(* Logix 5000 project; controller R400_500_XLS vendor 1 type 14 code 216 rev 31.11; software revision 31.01; part 21 of 32 *)
(* tags used below, declared in another part *)
   Abort1 : DINT;   // Not Used
   Alarm : SINT;   // Wait 3 seconds
   AlarmAcked : BOOL;   // Alarm has been acked
   bAlrm : BOOL[64];
   CycExcBuffer : UDT_CYCLE;
   F1rinse : DINT;   // Not Used
   F3rinse : DINT;   // Not Used
   H0_Temp : REAL;
   H1_Temp : REAL;
   HDelta_T : REAL;
   HeatSmp : DINT;
   iBuffer : DINT[5];
   Inj_Cond : SINT;   // Conductivity injection based steps
   Last_Hdelta_T : REAL;
   M : DINT[5];   // Memory Bits
   ONS_FC01 : DINT;
   ONS_FC12 : DINT;
   PresetMin : SINT;
   PresetSec : SINT;
   PreWtrDrnTme : DINT;
   PwExcBuffer : UDT_PW;
   PWR_UP : DINT;
   rBuffer : REAL[4];
   RecircLowHysteresis : REAL;
   RinseExcBuffer : UDT_RINSE;
   Run : DINT;
   SmpDrnTme : DINT;
   SmpHeatingSp : REAL;
   SmpLowHysteresis : REAL;
   StartPump3 : BOOL;   // Main Pump running
   Tmr : TIMER[107];
   TrecircSec : DINT;
   Trt_PrWsh : DINT;
   Trt_Rinse : DINT;   // Rinse steps
   washerMode : SINT;   // Washer Mode Flag 0 -> Ready; 1 -> Supervisor; 2 -> Service; 3 -> Run.
   WSH56_StartHeating : BOOL;   // Start heating
   WSH56_StartRecirculation : BOOL;   // Start the recirculation
   WshExcBuffer : UDT_WASH;
   Cfg_10_Modules : BOOL;   // Chassis is configured 10 slots
   Cfg_11_Modules : BOOL;
   Ctrlr_Status : DINT;
   Current_Screen : DINT;
   I_Ld_Dr_Cls_Sw : BOOL;   // Load door close
   I_MCR : BOOL;   // MCR input
   I_Pw_Tnk_Lvl_Sw : BOOL;   // Pure water tank level switch
   I_Smp_Lvl_Hgh : BOOL;   // Sump high level switch
   I_Smp_Lvl_Lw : BOOL;   // Sump low level switch
   I_Unld_Dr_Cls_Sw : BOOL;   // Unload door close
   MaintainCloseLd : BOOL;
   MaintainCloseUnld : BOOL;
   msg : BOOL[512];
   Msg_PwrUp : DINT;
   s007 : DINT;
   Screen_Ctrl : DINT;   // PLC Screen Request
   SumpHeatAlmRate : REAL;
   SumpTemp : REAL;   // Sump temperature in °C
   Unit : Hrdwre;   // Unit Configuration
(* MainProgram, continued *)

ROUTINE WSH_12_PWR_UP   (* ladder *)
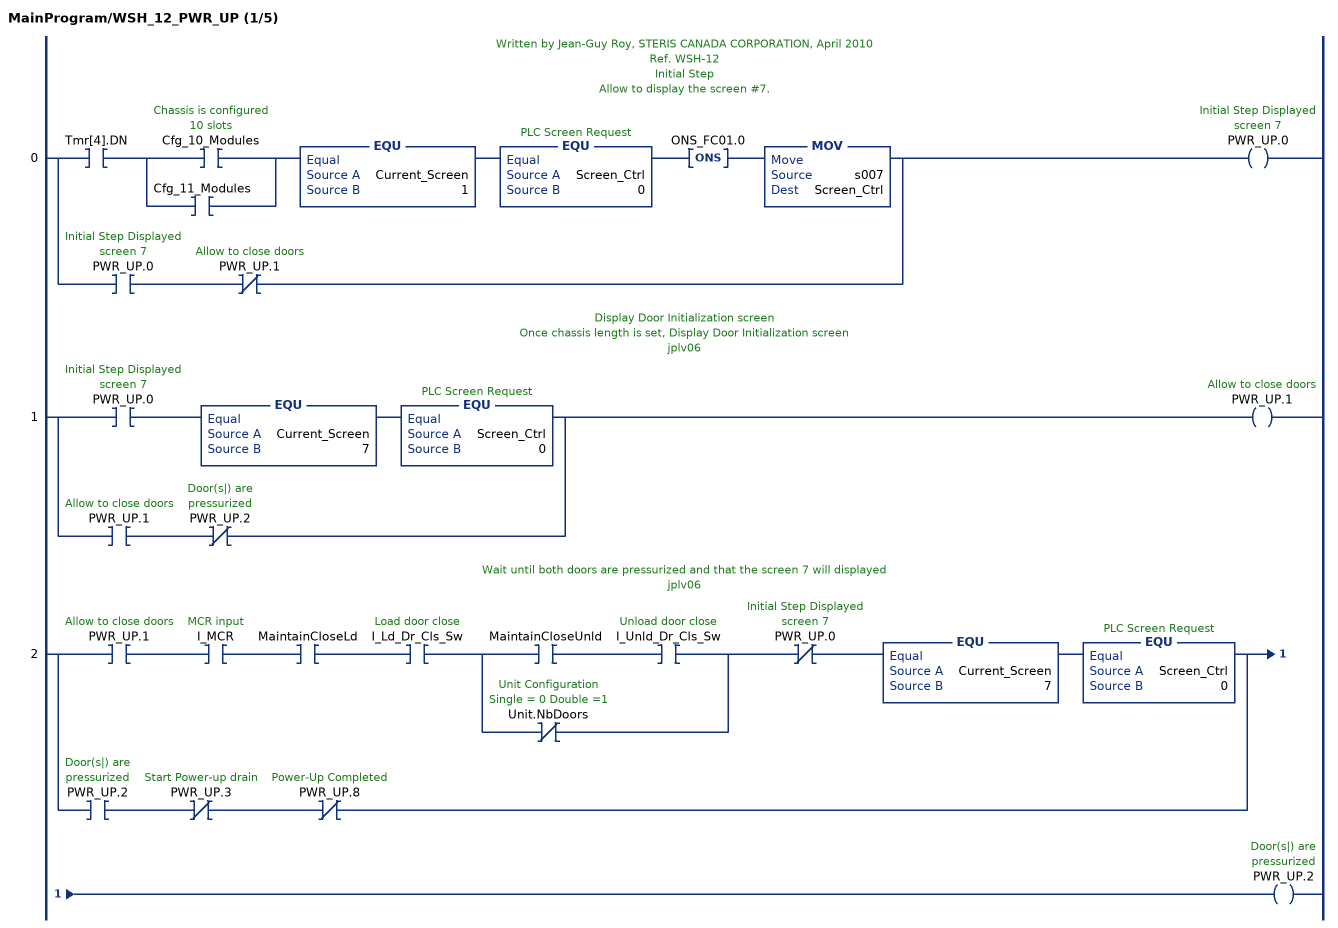
   // Written by Jean-Guy Roy, STERIS CANADA CORPORATION, April 2010
   // Ref. WSH-12
   // Initial Step
   // Allow to display the screen #7.
   0: [XIC(Tmr[4].DN) [XIC(Cfg_10_Modules) ,XIC(Cfg_11_Modules) ] EQU(Current_Screen,1) EQU(Screen_Ctrl,0) ONS(ONS_FC01.0) MOV(s007,Screen_Ctrl) ,XIC(PWR_UP.0) XIO(PWR_UP.1) ]OTE(PWR_UP.0);
   // Display Door Initialization screen
   // Once chassis length is set, Display Door Initialization screen
   // jplv06
   1: [XIC(PWR_UP.0) EQU(Current_Screen,7) EQU(Screen_Ctrl,0) ,XIC(PWR_UP.1) XIO(PWR_UP.2) ]OTE(PWR_UP.1);
   // Wait until both doors are pressurized and that the screen 7 will displayed
   // jplv06
   2: [XIC(PWR_UP.1) XIC(I_MCR) XIC(MaintainCloseLd) XIC(I_Ld_Dr_Cls_Sw) [XIC(MaintainCloseUnld) XIC(I_Unld_Dr_Cls_Sw) ,XIO(Unit.NbDoors) ] XIO(PWR_UP.0) EQU(Current_Screen,7) EQU(Screen_Ctrl,0) ,XIC(PWR_UP.2) XIO(PWR_UP.3) XIO(PWR_UP.8) ]OTE(PWR_UP.2);
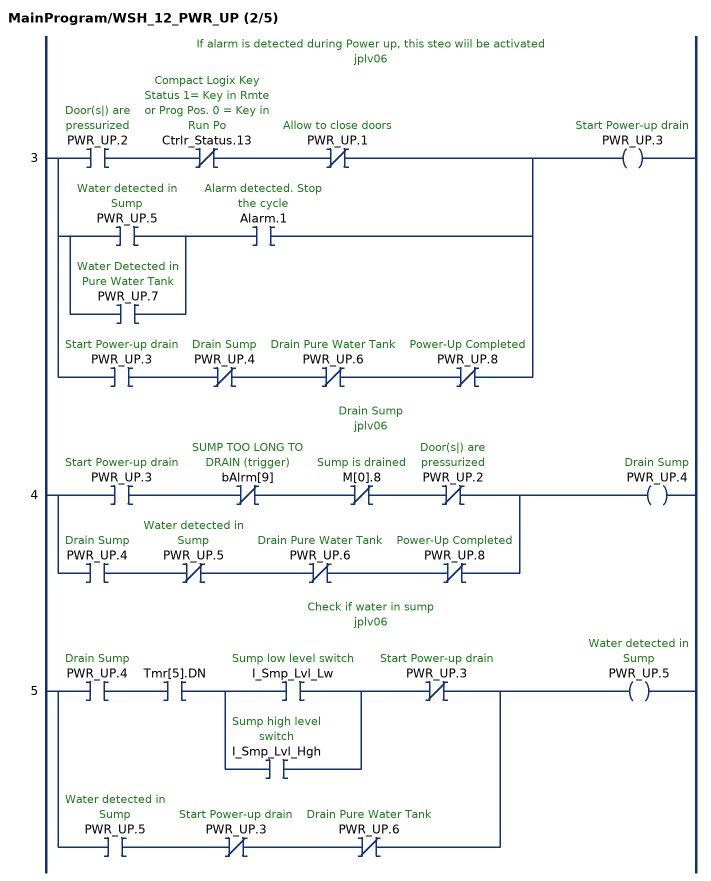
   // If alarm is detected during Power up, this steo wiil be activated
   // jplv06
   3: [XIC(PWR_UP.2) XIO(Ctrlr_Status.13) XIO(PWR_UP.1) ,[XIC(PWR_UP.5) ,XIC(PWR_UP.7) ] XIC(Alarm.1) ,XIC(PWR_UP.3) XIO(PWR_UP.4) XIO(PWR_UP.6) XIO(PWR_UP.8) ]OTE(PWR_UP.3);
   // Drain Sump
   // jplv06
   4: [XIC(PWR_UP.3) XIO(bAlrm[9]) XIO(M[0].8) XIO(PWR_UP.2) ,XIC(PWR_UP.4) XIO(PWR_UP.5) XIO(PWR_UP.6) XIO(PWR_UP.8) ]OTE(PWR_UP.4);
   // Check if water in sump
   // jplv06
   5: [XIC(PWR_UP.4) XIC(Tmr[5].DN) [XIC(I_Smp_Lvl_Lw) ,XIC(I_Smp_Lvl_Hgh) ] XIO(PWR_UP.3) ,XIC(PWR_UP.5) XIO(PWR_UP.3) XIO(PWR_UP.6) ]OTE(PWR_UP.5);
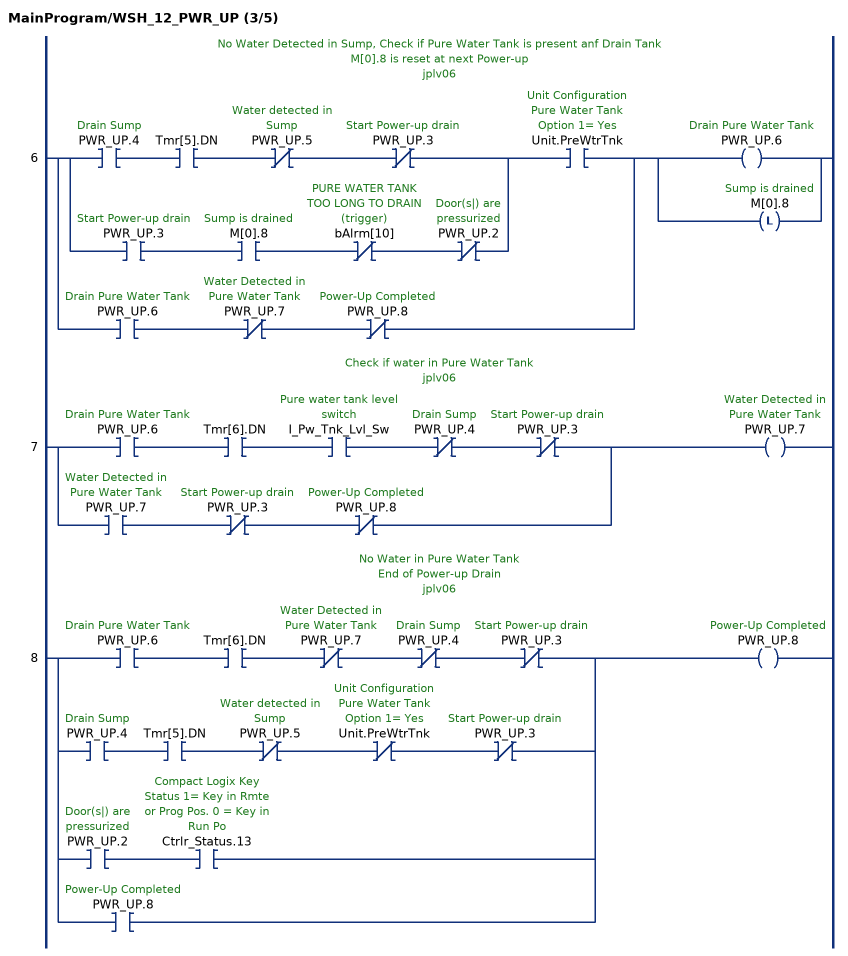
   // No Water Detected in Sump, Check if Pure Water Tank is present anf Drain Tank
   // M[0].8 is reset at next Power-up
   // jplv06
   6: [[XIC(PWR_UP.4) XIC(Tmr[5].DN) XIO(PWR_UP.5) XIO(PWR_UP.3) ,XIC(PWR_UP.3) XIC(M[0].8) XIO(bAlrm[10]) XIO(PWR_UP.2) ] XIC(Unit.PreWtrTnk) ,XIC(PWR_UP.6) XIO(PWR_UP.7) XIO(PWR_UP.8) ][OTE(PWR_UP.6) ,OTL(M[0].8) ];
   // Check if water in Pure Water Tank
   // jplv06
   7: [XIC(PWR_UP.6) XIC(Tmr[6].DN) XIC(I_Pw_Tnk_Lvl_Sw) XIO(PWR_UP.4) XIO(PWR_UP.3) ,XIC(PWR_UP.7) XIO(PWR_UP.3) XIO(PWR_UP.8) ]OTE(PWR_UP.7);
   // No Water in Pure Water Tank
   // End of Power-up Drain
   // jplv06
   8: [[XIC(PWR_UP.6) XIC(Tmr[6].DN) XIO(PWR_UP.7) XIO(PWR_UP.4) XIO(PWR_UP.3) ,XIC(PWR_UP.4) XIC(Tmr[5].DN) XIO(PWR_UP.5) XIO(Unit.PreWtrTnk) XIO(PWR_UP.3) ,XIC(PWR_UP.2) XIC(Ctrlr_Status.13) ] ,XIC(PWR_UP.8) ]OTE(PWR_UP.8);
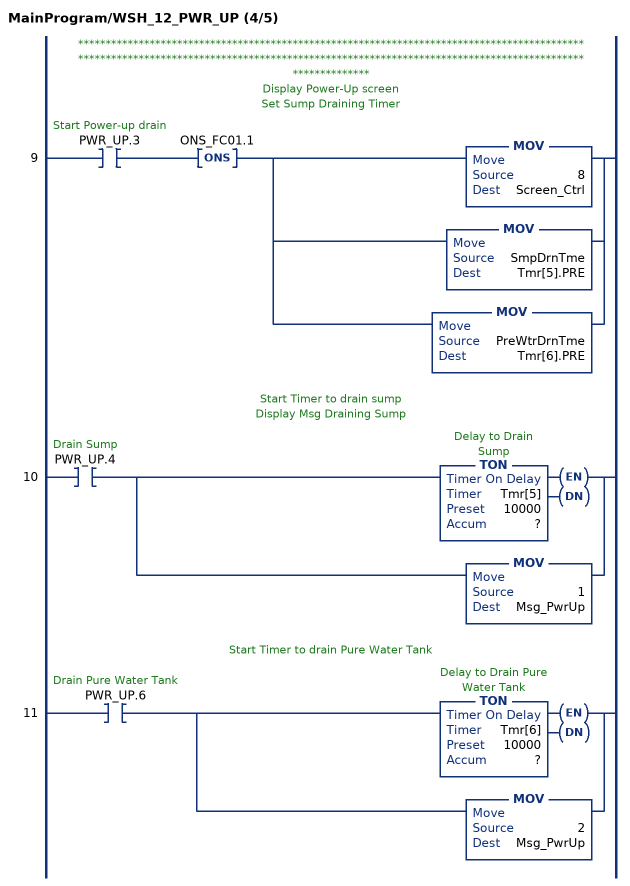
   // ******************************************************************************************************************************************************************************************************
   // Display Power-Up screen
   // Set Sump Draining Timer
   9: XIC(PWR_UP.3)ONS(ONS_FC01.1)[MOV(8,Screen_Ctrl) ,MOV(SmpDrnTme,Tmr[5].PRE) ,MOV(PreWtrDrnTme,Tmr[6].PRE) ];
   // Start Timer to drain sump
   // Display Msg Draining Sump
   10: XIC(PWR_UP.4)[TON(Tmr[5],?,?) ,MOV(1,Msg_PwrUp) ];
   // Start Timer to drain Pure Water Tank
   11: XIC(PWR_UP.6)[TON(Tmr[6],?,?) ,MOV(2,Msg_PwrUp) ];
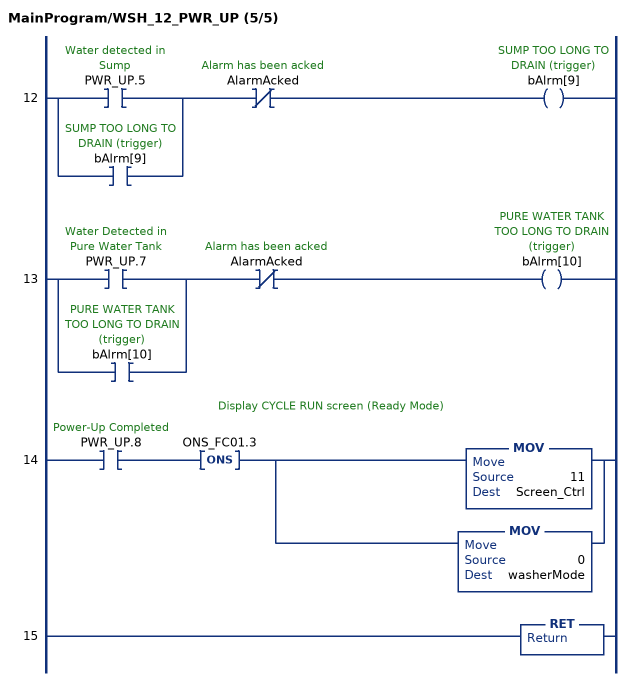
   12: [XIC(PWR_UP.5) ,XIC(bAlrm[9]) ]XIO(AlarmAcked)OTE(bAlrm[9]);
   13: [XIC(PWR_UP.7) ,XIC(bAlrm[10]) ]XIO(AlarmAcked)OTE(bAlrm[10]);
   // Display CYCLE RUN screen (Ready Mode)
   14: XIC(PWR_UP.8)ONS(ONS_FC01.3)[MOV(11,Screen_Ctrl) ,MOV(0,washerMode) ];
   15: RET();
END_ROUTINE

ROUTINE WSH_15_WSH_31_RECIRC_HEAT_SUMP   (* ladder *)
// This module is to heat the sump and the control of the recirculation timer
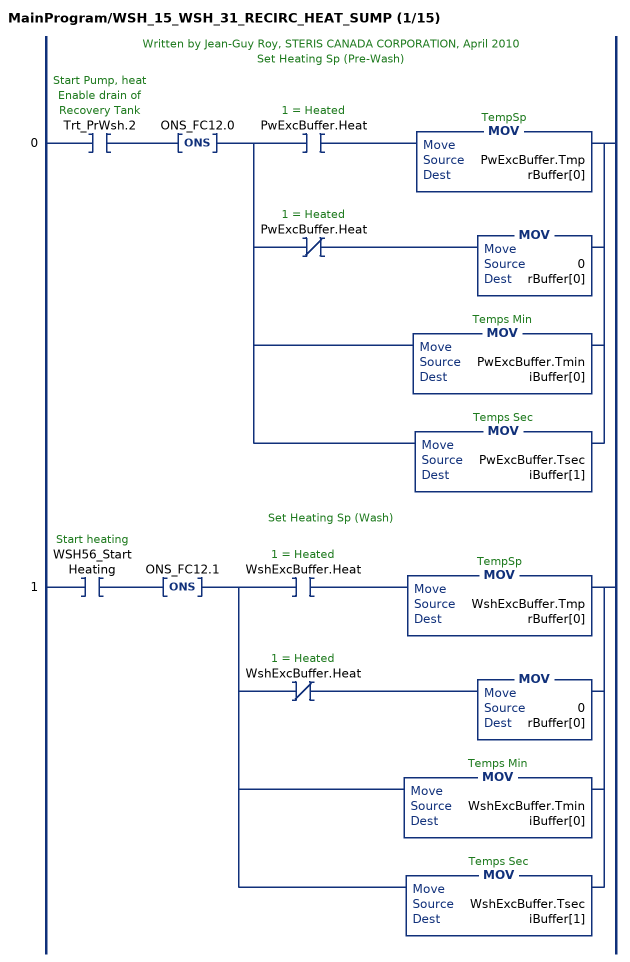
   // Written by Jean-Guy Roy, STERIS CANADA CORPORATION, April 2010
   // Set Heating Sp (Pre-Wash)
   0: XIC(Trt_PrWsh.2)ONS(ONS_FC12.0)[XIC(PwExcBuffer.Heat) MOV(PwExcBuffer.Tmp,rBuffer[0]) ,XIO(PwExcBuffer.Heat) MOV(0,rBuffer[0]) ,MOV(PwExcBuffer.Tmin,iBuffer[0]) ,MOV(PwExcBuffer.Tsec,iBuffer[1]) ];
   // Set Heating Sp (Wash)
   1: XIC(WSH56_StartHeating)ONS(ONS_FC12.1)[XIC(WshExcBuffer.Heat) MOV(WshExcBuffer.Tmp,rBuffer[0]) ,XIO(WshExcBuffer.Heat) MOV(0,rBuffer[0]) ,MOV(WshExcBuffer.Tmin,iBuffer[0]) ,MOV(WshExcBuffer.Tsec,iBuffer[1]) ];
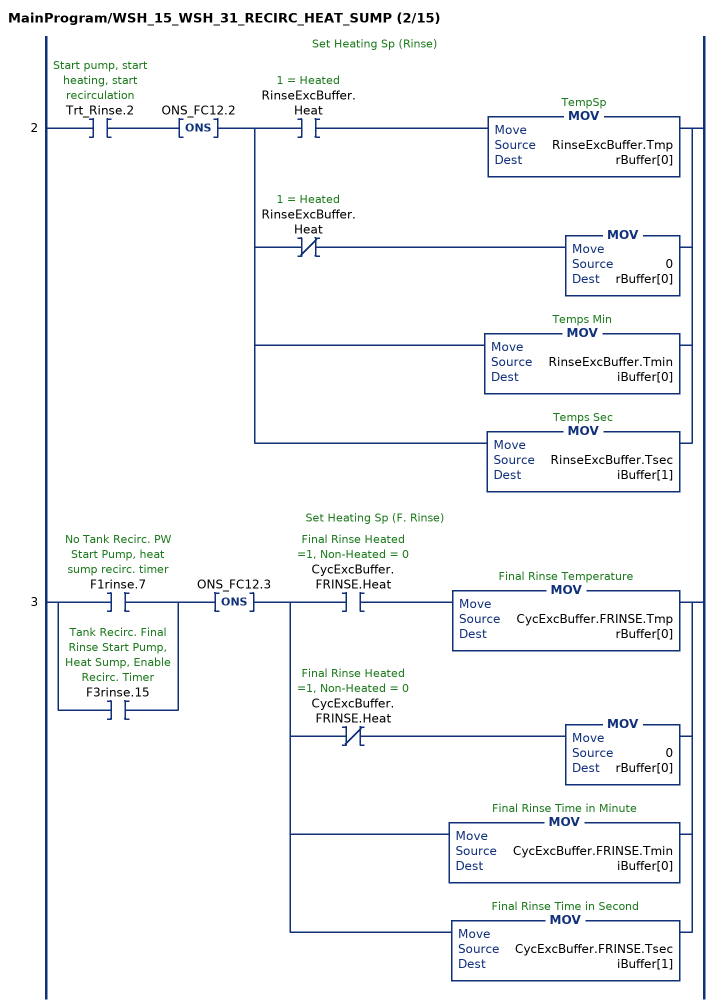
   // Set Heating Sp (Rinse)
   2: XIC(Trt_Rinse.2)ONS(ONS_FC12.2)[XIC(RinseExcBuffer.Heat) MOV(RinseExcBuffer.Tmp,rBuffer[0]) ,XIO(RinseExcBuffer.Heat) MOV(0,rBuffer[0]) ,MOV(RinseExcBuffer.Tmin,iBuffer[0]) ,MOV(RinseExcBuffer.Tsec,iBuffer[1]) ];
   // Set Heating Sp (F. Rinse)
   3: [XIC(F1rinse.7) ,XIC(F3rinse.15) ]ONS(ONS_FC12.3)[XIC(CycExcBuffer.FRINSE.Heat) MOV(CycExcBuffer.FRINSE.Tmp,rBuffer[0]) ,XIO(CycExcBuffer.FRINSE.Heat) MOV(0,rBuffer[0]) ,MOV(CycExcBuffer.FRINSE.Tmin,iBuffer[0]) ,MOV(CycExcBuffer.FRINSE.Tsec,iBuffer[1]) ];
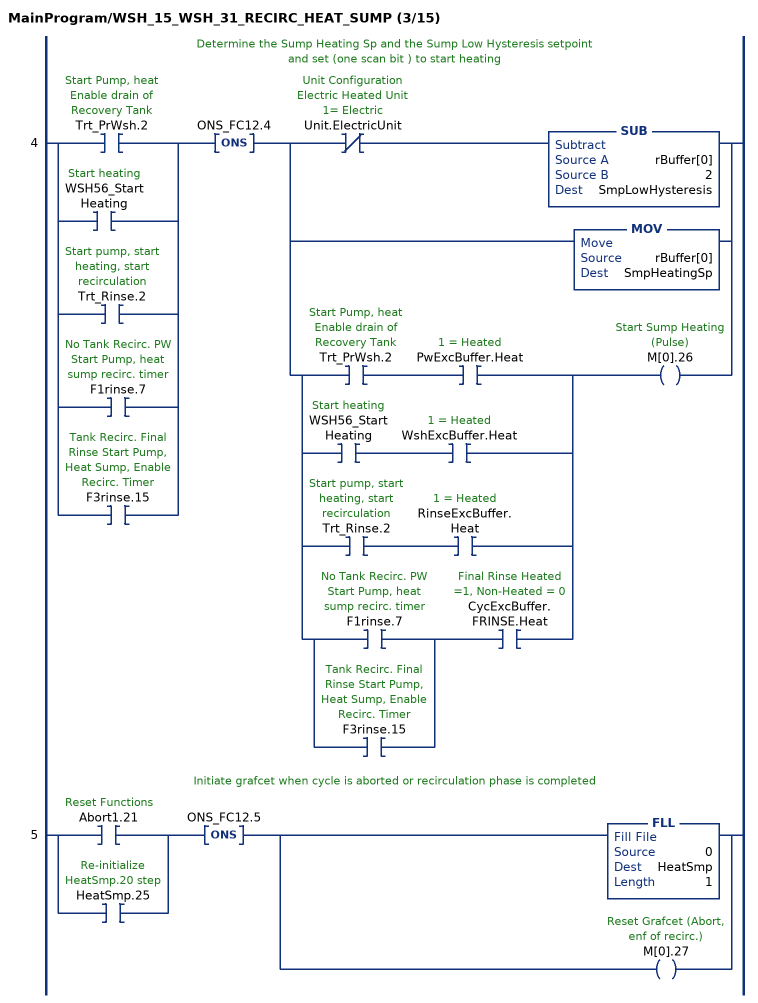
   // Determine the Sump Heating Sp and the Sump Low Hysteresis setpoint
   // and set (one scan bit ) to start heating
   4: [XIC(Trt_PrWsh.2) ,XIC(WSH56_StartHeating) ,XIC(Trt_Rinse.2) ,XIC(F1rinse.7) ,XIC(F3rinse.15) ]ONS(ONS_FC12.4)[XIO(Unit.ElectricUnit) SUB(rBuffer[0],2,SmpLowHysteresis) ,MOV(rBuffer[0],SmpHeatingSp) ,[XIC(Trt_PrWsh.2) XIC(PwExcBuffer.Heat) ,XIC(WSH56_StartHeating) XIC(WshExcBuffer.Heat) ,XIC(Trt_Rinse.2) XIC(RinseExcBuffer.Heat) ,[XIC(F1rinse.7) ,XIC(F3rinse.15) ] XIC(CycExcBuffer.FRINSE.Heat) ] OTE(M[0].26) ];
   // Initiate grafcet when cycle is aborted or recirculation phase is completed
   5: [XIC(Abort1.21) ,XIC(HeatSmp.25) ]ONS(ONS_FC12.5)[FLL(0,HeatSmp,1) ,OTE(M[0].27) ];
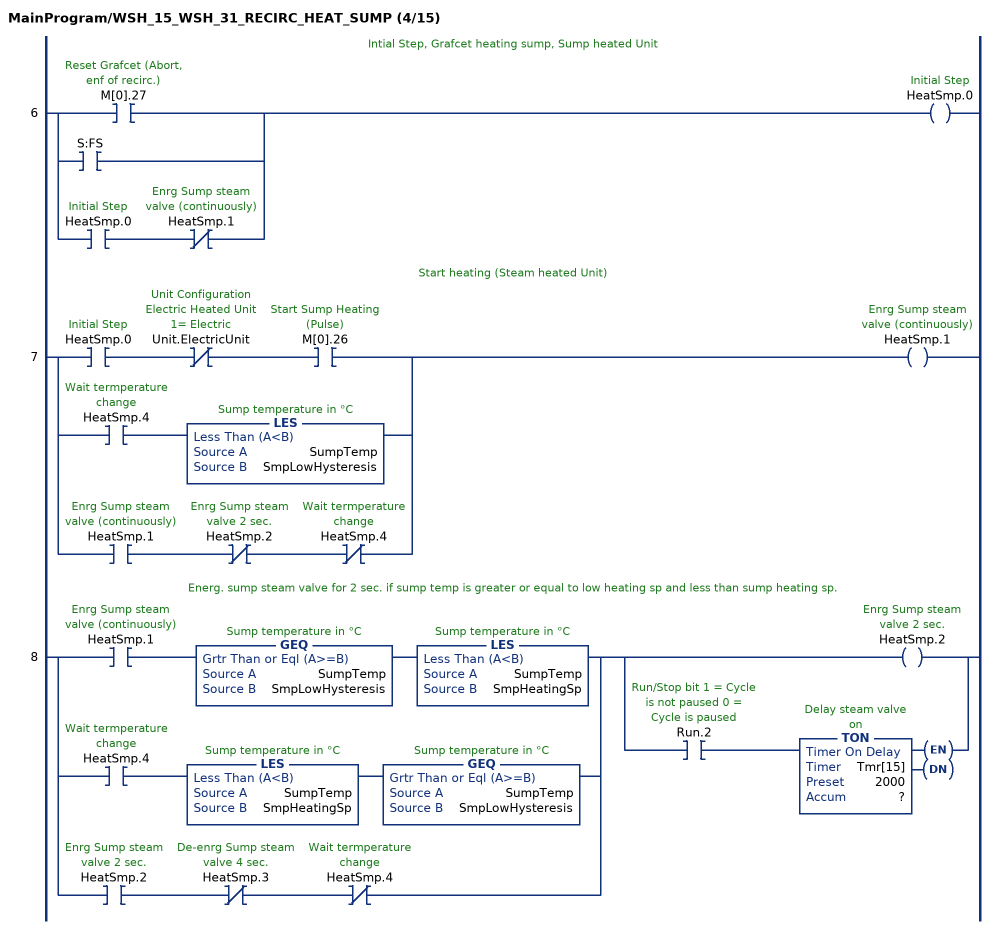
   // Intial Step, Grafcet heating sump, Sump heated Unit
   6: [XIC(M[0].27) ,XIC(S:FS) ,XIC(HeatSmp.0) XIO(HeatSmp.1) ]OTE(HeatSmp.0);
   // Start heating (Steam heated Unit)
   7: [XIC(HeatSmp.0) XIO(Unit.ElectricUnit) XIC(M[0].26) ,XIC(HeatSmp.4) LES(SumpTemp,SmpLowHysteresis) ,XIC(HeatSmp.1) XIO(HeatSmp.2) XIO(HeatSmp.4) ]OTE(HeatSmp.1);
   // Energ. sump steam valve for 2 sec. if sump temp is greater or equal to low heating sp and less than sump heating sp.
   8: [XIC(HeatSmp.1) GEQ(SumpTemp,SmpLowHysteresis) LES(SumpTemp,SmpHeatingSp) ,XIC(HeatSmp.4) LES(SumpTemp,SmpHeatingSp) GEQ(SumpTemp,SmpLowHysteresis) ,XIC(HeatSmp.2) XIO(HeatSmp.3) XIO(HeatSmp.4) ][OTE(HeatSmp.2) ,XIC(Run.2) TON(Tmr[15],?,?) ];
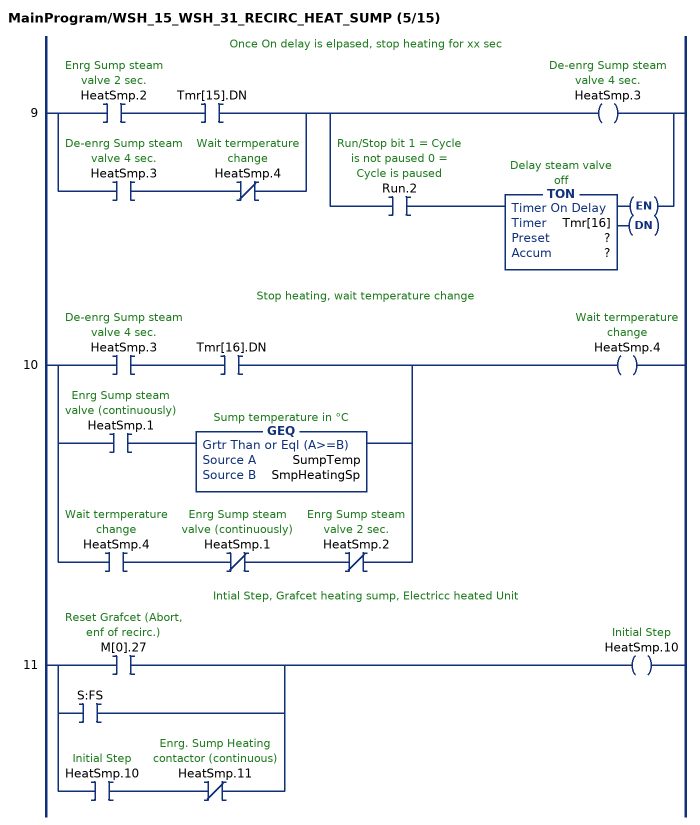
   // Once On delay is elpased, stop heating for xx sec
   9: [XIC(HeatSmp.2) XIC(Tmr[15].DN) ,XIC(HeatSmp.3) XIO(HeatSmp.4) ][OTE(HeatSmp.3) ,XIC(Run.2) TON(Tmr[16],?,?) ];
   // Stop heating, wait temperature change
   10: [XIC(HeatSmp.3) XIC(Tmr[16].DN) ,XIC(HeatSmp.1) GEQ(SumpTemp,SmpHeatingSp) ,XIC(HeatSmp.4) XIO(HeatSmp.1) XIO(HeatSmp.2) ]OTE(HeatSmp.4);
   // Intial Step, Grafcet heating sump, Electricc heated Unit
   11: [XIC(M[0].27) ,XIC(S:FS) ,XIC(HeatSmp.10) XIO(HeatSmp.11) ]OTE(HeatSmp.10);
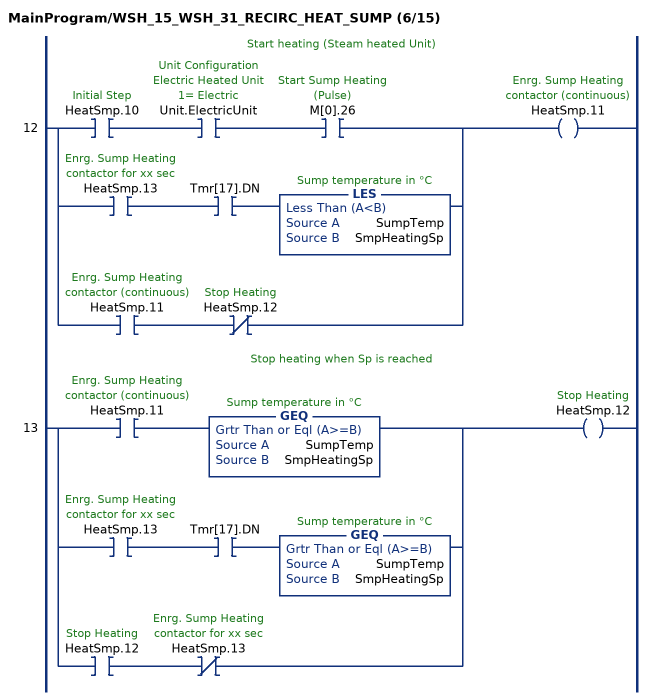
   // Start heating (Steam heated Unit)
   12: [XIC(HeatSmp.10) XIC(Unit.ElectricUnit) XIC(M[0].26) ,XIC(HeatSmp.13) XIC(Tmr[17].DN) LES(SumpTemp,SmpHeatingSp) ,XIC(HeatSmp.11) XIO(HeatSmp.12) ]OTE(HeatSmp.11);
   // Stop heating when Sp is reached
   13: [XIC(HeatSmp.11) GEQ(SumpTemp,SmpHeatingSp) ,XIC(HeatSmp.13) XIC(Tmr[17].DN) GEQ(SumpTemp,SmpHeatingSp) ,XIC(HeatSmp.12) XIO(HeatSmp.13) ]OTE(HeatSmp.12);
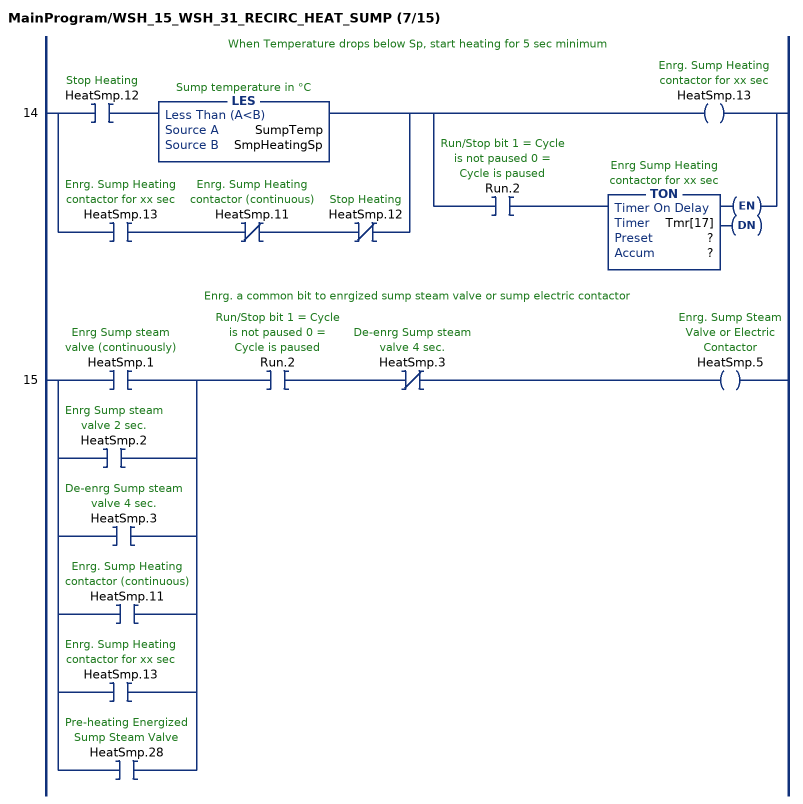
   // When Temperature drops below Sp, start heating for 5 sec minimum
   14: [XIC(HeatSmp.12) LES(SumpTemp,SmpHeatingSp) ,XIC(HeatSmp.13) XIO(HeatSmp.11) XIO(HeatSmp.12) ][OTE(HeatSmp.13) ,XIC(Run.2) TON(Tmr[17],?,?) ];
   // Enrg. a common bit to enrgized sump steam valve or sump electric contactor
   15: [XIC(HeatSmp.1) ,XIC(HeatSmp.2) ,XIC(HeatSmp.3) ,XIC(HeatSmp.11) ,XIC(HeatSmp.13) ,XIC(HeatSmp.28) ]XIC(Run.2)XIO(HeatSmp.3)OTE(HeatSmp.5);
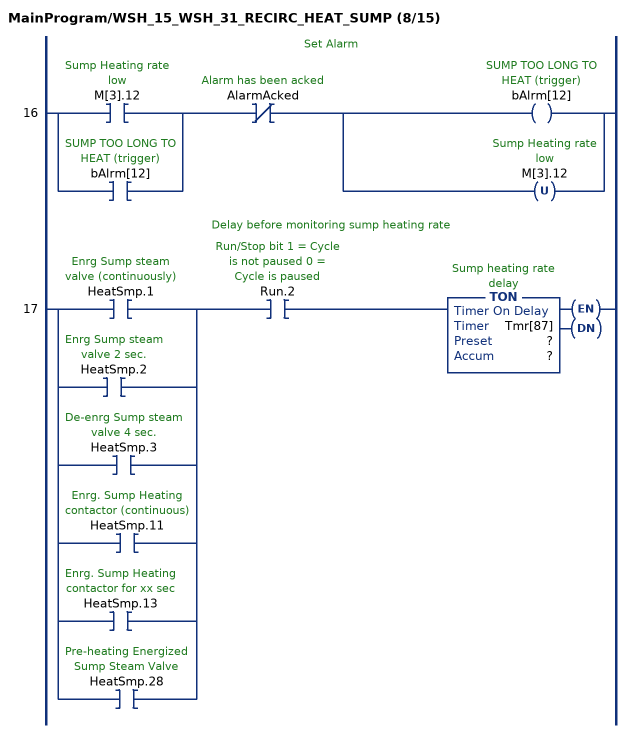
   // Set Alarm
   16: [XIC(M[3].12) ,XIC(bAlrm[12]) ]XIO(AlarmAcked)[OTE(bAlrm[12]) ,OTU(M[3].12) ];
   // Delay before monitoring sump heating rate
   17: [XIC(HeatSmp.1) ,XIC(HeatSmp.2) ,XIC(HeatSmp.3) ,XIC(HeatSmp.11) ,XIC(HeatSmp.13) ,XIC(HeatSmp.28) ]XIC(Run.2)TON(Tmr[87],?,?);
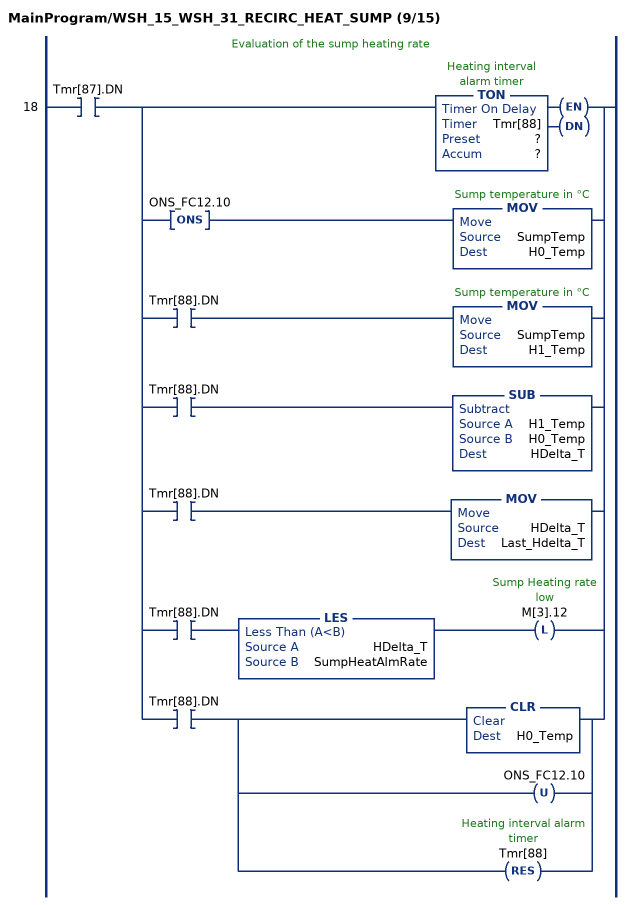
   // Evaluation of the sump heating rate
   18: XIC(Tmr[87].DN)[TON(Tmr[88],?,?) ,ONS(ONS_FC12.10) MOV(SumpTemp,H0_Temp) ,XIC(Tmr[88].DN) MOV(SumpTemp,H1_Temp) ,XIC(Tmr[88].DN) SUB(H1_Temp,H0_Temp,HDelta_T) ,XIC(Tmr[88].DN) MOV(HDelta_T,Last_Hdelta_T) ,XIC(Tmr[88].DN) LES(HDelta_T,SumpHeatAlmRate) OTL(M[3].12) ,XIC(Tmr[88].DN) [CLR(H0_Temp) ,OTU(ONS_FC12.10) ,RES(Tmr[88]) ] ];
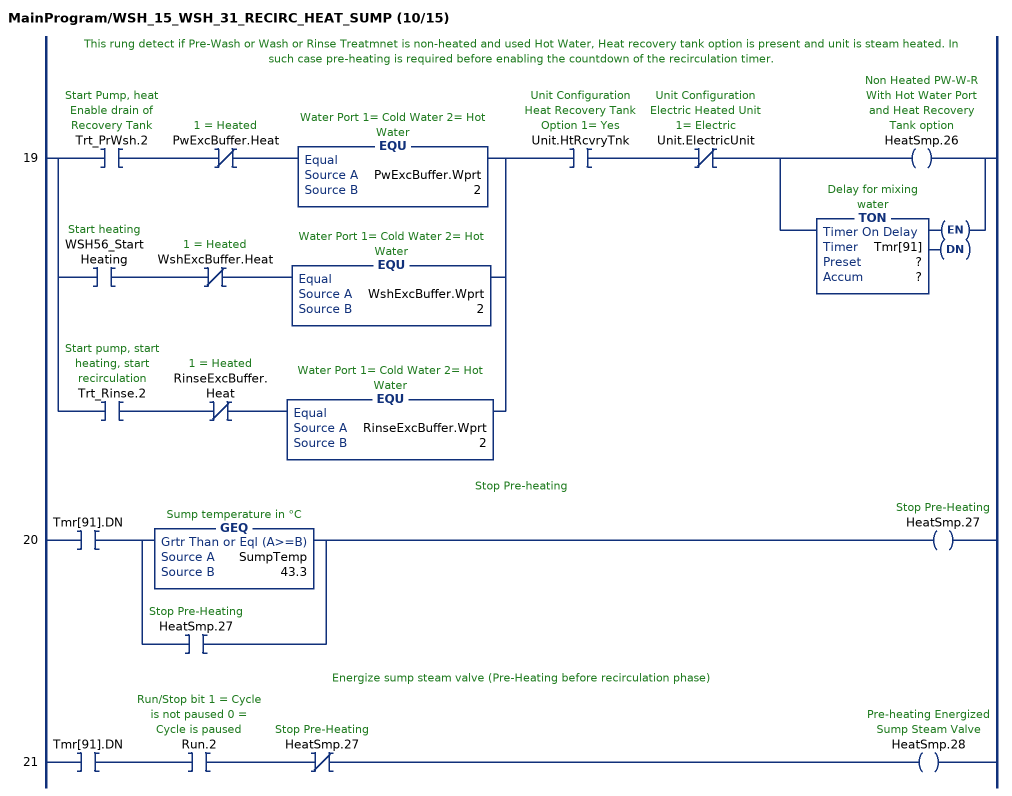
   // This rung detect if Pre-Wash or Wash or Rinse Treatmnet is non-heated and used Hot Water, Heat recovery tank option is present and unit is steam heated. In such case pre-heating is required before enabling the countdown of the recirculation timer.
   19: [XIC(Trt_PrWsh.2) XIO(PwExcBuffer.Heat) EQU(PwExcBuffer.Wprt,2) ,XIC(WSH56_StartHeating) XIO(WshExcBuffer.Heat) EQU(WshExcBuffer.Wprt,2) ,XIC(Trt_Rinse.2) XIO(RinseExcBuffer.Heat) EQU(RinseExcBuffer.Wprt,2) ]XIC(Unit.HtRcvryTnk)XIO(Unit.ElectricUnit)[OTE(HeatSmp.26) ,TON(Tmr[91],?,?) ];
   // Stop Pre-heating
   20: XIC(Tmr[91].DN)[GEQ(SumpTemp,43.3) ,XIC(HeatSmp.27) ]OTE(HeatSmp.27);
   // Energize sump steam valve (Pre-Heating before recirculation phase)
   21: XIC(Tmr[91].DN)XIC(Run.2)XIO(HeatSmp.27)OTE(HeatSmp.28);
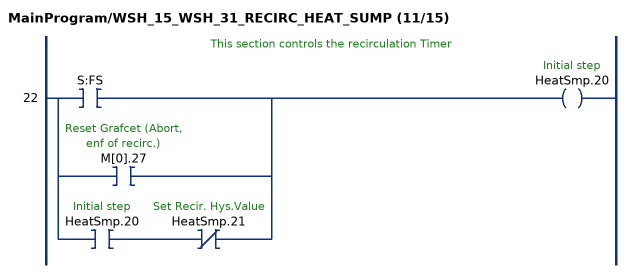
   // This section controls the recirculation Timer
   22: [XIC(S:FS) ,XIC(M[0].27) ,XIC(HeatSmp.20) XIO(HeatSmp.21) ]OTE(HeatSmp.20);
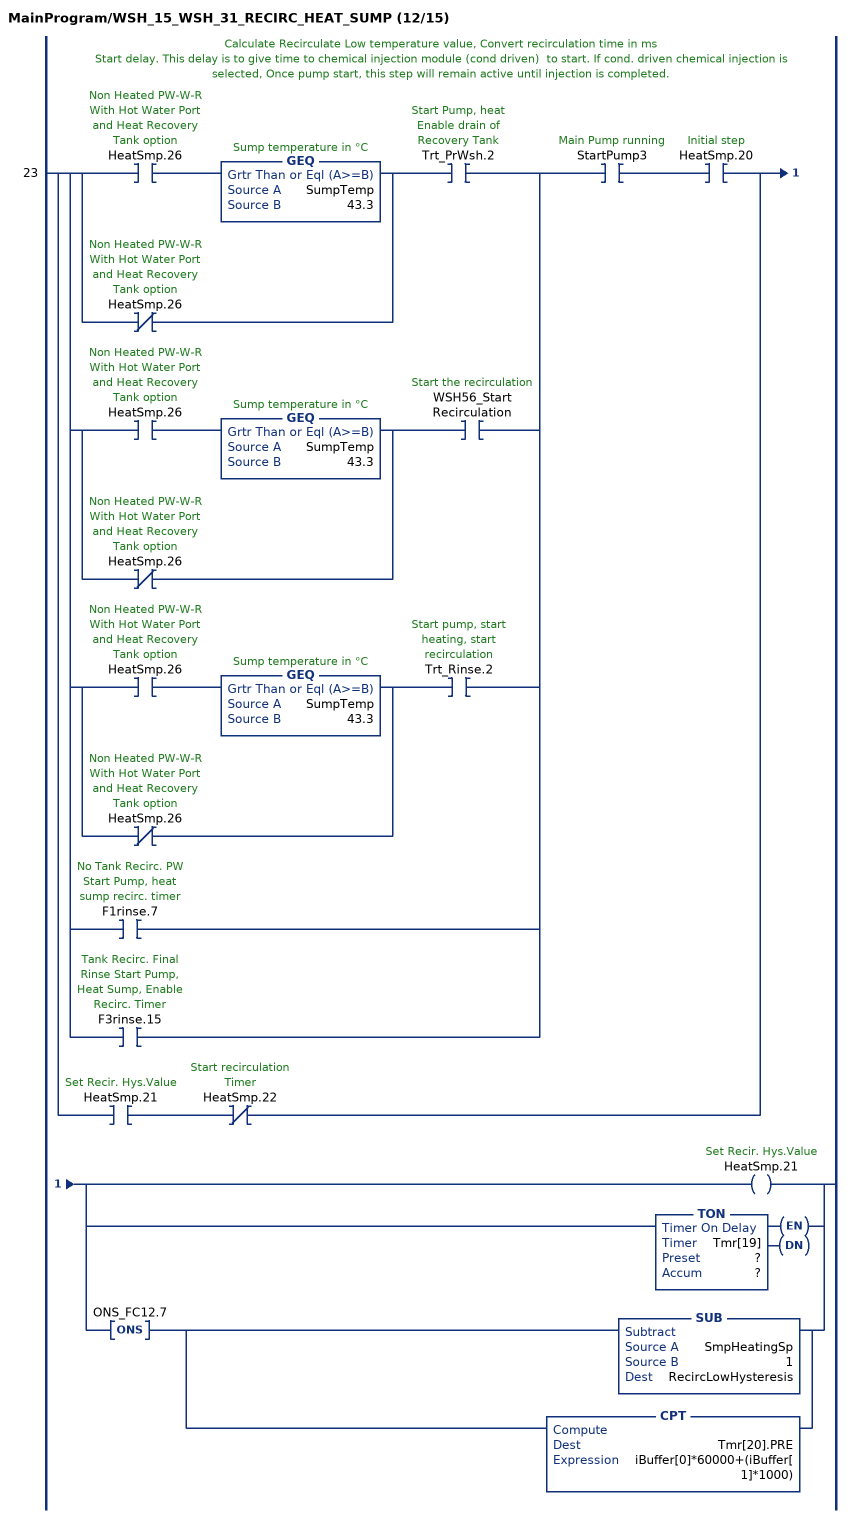
   // Calculate Recirculate Low temperature value, Convert recirculation time in ms
   // Start delay. This delay is to give time to chemical injection module (cond driven)  to start. If cond. driven chemical injection is selected, Once pump start, this step will remain active until injection is completed.
   23: [[[XIC(HeatSmp.26) GEQ(SumpTemp,43.3) ,XIO(HeatSmp.26) ] XIC(Trt_PrWsh.2) ,[XIC(HeatSmp.26) GEQ(SumpTemp,43.3) ,XIO(HeatSmp.26) ] XIC(WSH56_StartRecirculation) ,[XIC(HeatSmp.26) GEQ(SumpTemp,43.3) ,XIO(HeatSmp.26) ] XIC(Trt_Rinse.2) ,XIC(F1rinse.7) ,XIC(F3rinse.15) ] XIC(StartPump3) XIC(HeatSmp.20) ,XIC(HeatSmp.21) XIO(HeatSmp.22) ][OTE(HeatSmp.21) ,TON(Tmr[19],?,?) ,ONS(ONS_FC12.7) [SUB(SmpHeatingSp,1,RecircLowHysteresis) ,CPT(Tmr[20].PRE,iBuffer[0]*60000+(iBuffer[1]*1000)) ] ];
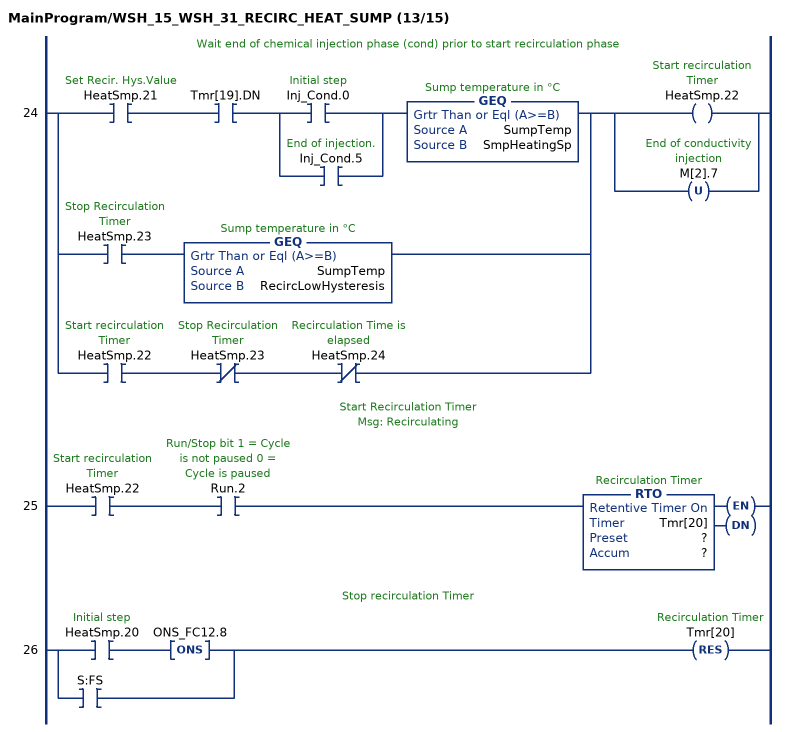
   // Wait end of chemical injection phase (cond) prior to start recirculation phase
   24: [XIC(HeatSmp.21) XIC(Tmr[19].DN) [XIC(Inj_Cond.0) ,XIC(Inj_Cond.5) ] GEQ(SumpTemp,SmpHeatingSp) ,XIC(HeatSmp.23) GEQ(SumpTemp,RecircLowHysteresis) ,XIC(HeatSmp.22) XIO(HeatSmp.23) XIO(HeatSmp.24) ][OTE(HeatSmp.22) ,OTU(M[2].7) ];
   // Start Recirculation Timer
   // Msg: Recirculating
   25: XIC(HeatSmp.22)XIC(Run.2)RTO(Tmr[20],?,?);
   // Stop recirculation Timer
   26: [XIC(HeatSmp.20) ONS(ONS_FC12.8) ,XIC(S:FS) ]RES(Tmr[20]);
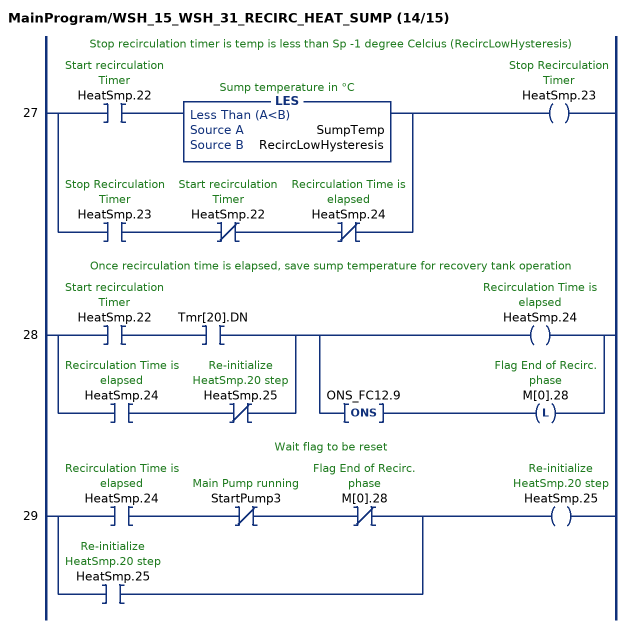
   // Stop recirculation timer is temp is less than Sp -1 degree Celcius (RecircLowHysteresis)
   27: [XIC(HeatSmp.22) LES(SumpTemp,RecircLowHysteresis) ,XIC(HeatSmp.23) XIO(HeatSmp.22) XIO(HeatSmp.24) ]OTE(HeatSmp.23);
   // Once recirculation time is elapsed, save sump temperature for recovery tank operation
   28: [XIC(HeatSmp.22) XIC(Tmr[20].DN) ,XIC(HeatSmp.24) XIO(HeatSmp.25) ][OTE(HeatSmp.24) ,ONS(ONS_FC12.9) OTL(M[0].28) ];
   // Wait flag to be reset
   29: [XIC(HeatSmp.24) XIO(StartPump3) XIO(M[0].28) ,XIC(HeatSmp.25) ]OTE(HeatSmp.25);
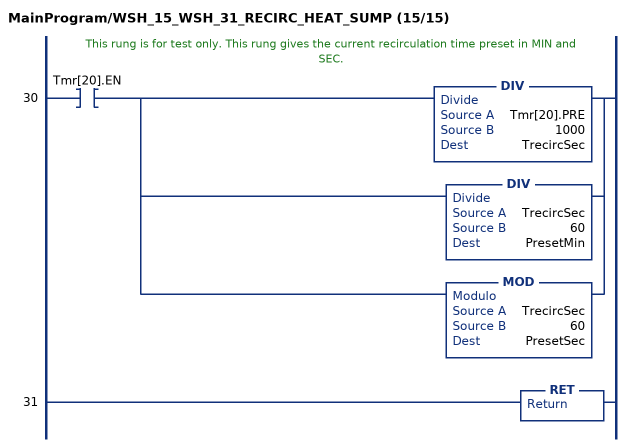
   // This rung is for test only. This rung gives the current recirculation time preset in MIN and SEC.
   30: XIC(Tmr[20].EN)[DIV(Tmr[20].PRE,1000,TrecircSec) ,DIV(TrecircSec,60,PresetMin) ,MOD(TrecircSec,60,PresetSec) ];
   31: RET();
END_ROUTINE
